Fanuc KAREL source: kt00991.KL

-- PROVISIONAL review KL for V770-1; original PC SHA256 39fd68e7ba532028a7bb77d833319e636cf694038469dae573d24b8312789f8e
-- Incomplete behavior may be omitted. Consult companion uncertainty JSON. Do not deploy.
PROGRAM KT00991
%NOLOCKGROUP
VAR
  X : REAL
  Y : REAL
  Z : REAL
  W : REAL
  P : REAL
  R : REAL
-- UNRESOLVED_DECL P1 type=000101
-- UNRESOLVED_DECL P2 type=000101
-- UNRESOLVED_DECL CFG type=00001c
BEGIN
  -- UNRESOLVED_PC offsets 5-65; opcodes 27,27,49,7E,AD,22,22,22,22,22,22,22,76
  -- UNRESOLVED_PC offsets 70-74; opcodes 7F
END KT00991
